INTERFACE I_Motor

METHOD Start : BOOL
VAR_INPUT
    fSpeed : LREAL;
END_VAR
END_METHOD

END_INTERFACE

(* stored: Version 1.1.0.1, ProductVersion 3.1.4024.12
   Itf I_Motor: Id {cccccccc-0000-0000-0000-000000000001}
   Method Start: Id {cccccccc-0000-0000-0000-000000000002} *)
